Staubli VAL3: removeActCmd.pgx

program removeActCmd(num x_nStackIndex)
begin
  actCmd[x_nStackIndex].nMoveID=-1
  actCmd[x_nStackIndex].nActionID=-1
  actCmd[x_nStackIndex].bActFinish[0]=false
end
